FUNCTION_BLOCK Tank (* Composite Function Block Type *)
  (* Standard: 61499-2 *)
  (* Version 0.0, 6/20/2016, Andrei, nxtControl GmbH, template *)
  PACKAGE Main;
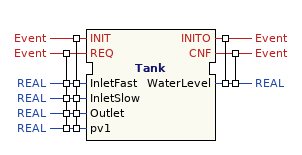
  EVENT_INPUT
    INIT WITH InletFast, InletSlow, Outlet, pv1; (* Initialization Request *)
    REQ WITH InletFast, InletSlow, Outlet, pv1; (* Normal Execution Request *)
  END_EVENT
  EVENT_OUTPUT
    INITO WITH WaterLevel; (* Initialization Confirm *)
    CNF WITH WaterLevel; (* Execution Confirmation *)
  END_EVENT
  VAR_INPUT
    InletFast : REAL; (* Input event qualifier *)
    InletSlow : REAL;
    Outlet : REAL;
    pv1 : REAL;
  END_VAR
  VAR_OUTPUT
    WaterLevel : REAL; (* Output event qualifier *)
  END_VAR
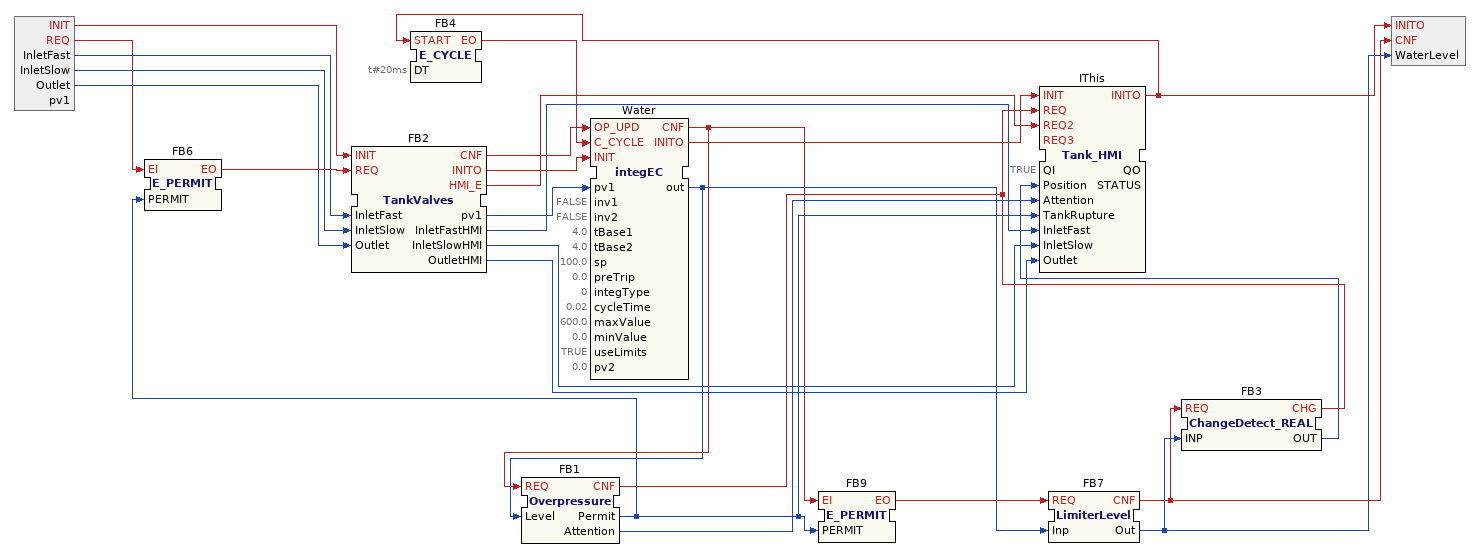
  FBS
    Water : integEC(inv1 := FALSE, inv2 := FALSE, tBase1 := 4.0, tBase2 := 4.0, sp := 100.0, preTrip := 0.0, integType := 0, cycleTime := 0.02, maxValue := 600.0, minValue := 0.0, useLimits := TRUE, pv2 := 0.0);
    FB3 : ChangeDetect_REAL;
    FB4 : E_CYCLE(DT := t#20ms);
    FB2 : TankValves;
    FB6 : E_PERMIT;
    IThis : Tank_HMI(QI := TRUE);
    FB9 : E_PERMIT;
    FB7 : LimiterLevel;
    FB1 : Overpressure;
  END_FBS
  EVENT_CONNECTIONS
    FB2.CNF TO Water.OP_UPD;
    INIT TO FB2.INIT;
    FB6.EO TO FB2.REQ;
    FB4.EO TO Water.C_CYCLE;
    FB2.INITO TO Water.INIT;
    Water.CNF TO FB1.REQ;
    REQ TO FB6.EI;
    Water.CNF TO FB9.EI;
    FB9.EO TO FB7.REQ;
    FB7.CNF TO FB3.REQ;
    FB7.CNF TO CNF;
    Water.INITO TO IThis.INIT;
    FB1.CNF TO IThis.REQ;
    FB3.CHG TO IThis.REQ;
    FB2.HMI_E TO IThis.REQ2;
    IThis.INITO TO FB4.START;
    IThis.INITO TO INITO;
  END_CONNECTIONS
  DATA_CONNECTIONS
    InletFast TO FB2.InletFast;
    InletSlow TO FB2.InletSlow;
    Outlet TO FB2.Outlet;
    Water.out TO FB1.Level;
    FB1.Permit TO FB9.PERMIT;
    Water.out TO FB7.Inp;
    FB1.Permit TO FB6.PERMIT;
    FB7.Out TO FB3.INP;
    FB7.Out TO WaterLevel;
    FB2.pv1 TO Water.pv1;
    FB3.OUT TO IThis.Position;
    FB1.Attention TO IThis.Attention;
    FB1.Permit TO IThis.TankRupture;
    FB2.InletFastHMI TO IThis.InletFast;
    FB2.InletSlowHMI TO IThis.InletSlow;
    FB2.OutletHMI TO IThis.Outlet;
  END_CONNECTIONS
END_FUNCTION_BLOCK
